(* IEC 61131-3 sources: JingjiangMoonbox/Application/Application/任务列表/TensionTask/张力控制/收放牵/其他, 4 files *)

(* ---- AntiNotch.st ---- *)
(*@CES
Name=AntiNotch
Type=FunctionBlock
TypeGuid=6f9dac99-8de1-4efc-8465-68ac443b7d08
Guid=24b15fba-c20e-4805-94ad-f0677bc5936e
HasDeclaration=True
HasImplementation=True
*)
{DECLARATION}
FUNCTION AntiNotch : BOOL
(*功能：反陷波器(s^2+2*d*wn*s+wn^2)/(s^2+2*d*xi*wn*s+wn^2)的差分方程实现*)
(*输入：*)
(*输出：*)
VAR_INPUT
	i_rU:REAL;(*信号输入*)
	i_prYout: POINTER TO REAL;(*信号输出*)

(*(s^2+2*d*wn*s+wn^2)/(s^2+2*d*xi*wn*s+wn^2)*)
	i_rWn:REAL;(*陷波中心频率 rad/s*)
	i_rBw:REAL;(*陷波宽度 rad/s*)
	i_rDp:REAL;(*陷波深度 dB*)

	i_rTs:REAL;(*采样时间*)

	i_prUk:POINTER TO ARRAY [1..3] OF REAL;(*输入寄存器*)
	i_prYk:POINTER TO ARRAY [1..3] OF REAL;(*输出寄存器*)
END_VAR
VAR
	rFn:REAL:=0;
	rFBw:REAL:=0;
	rWn:REAL:=0;
	rDp:REAL:=0;

	rD:REAL:=0;
	rXi:REAL:=0;

	rK:REAL:=0;
	ra2:REAL:=0;
	ra1:REAL:=0;
	ra0:REAL:=0;

	rb2:REAL:=0;
	rb1:REAL:=0;
	rb0:REAL:=0;

	rTs:REAL:=0;(*采样时间*)
	rTemp:REAL:=0;

END_VAR
{IMPLEMENTATION}
(*参数初始化*)
rFn := LREAL_TO_REAL(i_rWn/2.0*gc_lrPi);
rWn := i_rWn;
rFBw := LREAL_TO_REAL(i_rBw/2.0*gc_lrPi);
rDp := i_rDp;

rTemp := -rDp/20.0;
rD := LREAL_TO_REAL(EXPT(10,rTemp));

rTemp := LREAL_TO_REAL(1.0/(1.0 - 2.0*EXPT(rD,2)));
rXi := rFBw/(2.0*rFn)*SQRT(rTemp);

rK := 1.0;

ra2:=1.0;
ra1:=2*rXi*rWn;
ra0:=rWn*rWn;

rb2:=1;
rb1:=2*rD*rXi*rWn;
rb0:=rWn*rWn;

rTs:=i_rTs;

(*更新寄存器注意顺序*)
i_prYk^[3]:=i_prYk^[2];
i_prYk^[2]:=i_prYk^[1];

i_prUk^[3]:=i_prUk^[2];
i_prUk^[2]:=i_prUk^[1];

(*差分计算*)
i_prUk^[1]:=rK*i_rU;
rTemp:=1/(rb0*rTs*rTs+2*rb1*rTs+4*rb2)*(-(2*rb0*rTs*rTs-8*rb2)*i_prYk^[2]-(rb0*rTs*rTs-2*rb1*rTs+4*rb2)*i_prYk^[3]
            +(ra0*rTs*rTs+2*ra1*rTs+4*ra2)*i_prUk^[1]+(2*ra0*rTs*rTs-8*ra2)*i_prUk^[2]+(ra0*rTs*rTs-2*ra1*rTs+4*ra2)*i_prUk^[3]);
i_prYk^[1]:=rTemp;
i_prYout^:=rTemp;

(* ---- KS_A2B_SmoothDeal.st ---- *)
(*@CES
Name=KS_A2B_SmoothDeal
Type=FunctionBlock
TypeGuid=6f9dac99-8de1-4efc-8465-68ac443b7d08
Guid=9cfb7a1c-ce6a-4c3a-85a6-d0a941a33b90
HasDeclaration=True
HasImplementation=True
*)
{DECLARATION}
FUNCTION KS_A2B_SmoothDeal : REAL
(*从A变化到B平滑处理,返回当前值*)
VAR_INPUT
	i_rA:REAL;
	i_rB:REAL;
	i_rDelta:REAL;(*变化值*)
END_VAR
VAR
	rC:REAL;
END_VAR
{IMPLEMENTATION}
IF i_rDelta<>0 THEN
	IF i_rA > i_rB THEN
		rC:= i_rA - i_rDelta;
		IF rC < i_rB THEN(*限值处理*)
			rC:=i_rB;
		END_IF
	ELSIF i_rA < i_rB THEN
		rC:= i_rA + i_rDelta;
		IF rC > i_rB THEN(*限值处理*)
			rC:=i_rB;
		END_IF
	ELSE
		rC:= i_rB;
	END_IF
ELSE
	rC:=i_rB;
END_IF

KS_A2B_SmoothDeal:=rC;

(* ---- KS_SIG_SIN.st ---- *)
(*@CES
Name=KS_SIG_SIN
Type=FunctionBlock
TypeGuid=6f9dac99-8de1-4efc-8465-68ac443b7d08
Guid=c56967f0-af3c-4951-929b-0432ccffd3b8
HasDeclaration=True
HasImplementation=True
*)
{DECLARATION}
FUNCTION KS_SIG_SIN : BOOL
(*正弦信号*)
VAR_INPUT
	i_xEn:BOOL;(*使能*)
	i_rFreq:REAL;(*频率@hz*)
	i_rAmplitude:REAL;(*幅值*)
	i_uiTotalTime:UINT;(*输出的总时间|=0 代表一直输出@s*)
	i_iCycleTime_Plc:INT;(*程序时间@ms*)
	i_pxOuting:POINTER TO BOOL;(*输出中@如果取消使能,停止到0时结束*)
	i_plrX:POINTER TO LREAL;(*X轴的值*)
	i_prResult:POINTER TO REAL;(*结果值*)
END_VAR
VAR
	xOuting:BOOL;
	lrX:LREAL;(*x值*)
	rResult: REAL;
	lrW:LREAL;(*角速度@rad/s*)
	lrpi: LREAL := 3.1415926;(*圆周率*)
	lrTs: LREAL;(*周期@s*)
	lrTmp: LREAL;
	lrTotalTime:LREAL;(*输出的总时间@ms*)
	xStopOuting: BOOL;
END_VAR
{IMPLEMENTATION}
IF i_rFreq<>0 AND i_rAmplitude<>0 AND i_iCycleTime_Plc<>0 THEN;
ELSE
	RETURN;
END_IF

IF i_pxOuting<>0 THEN
	xOuting:=i_pxOuting^;
END_IF
IF i_plrX<>0 THEN
	lrX:=i_plrX^;
END_IF
IF i_prResult<>0 THEN
	rResult:=i_prResult^;
END_IF

(*使能*)
IF i_xEn THEN
	IF NOT xOuting AND
		lrX = 0 THEN(*lrx用来控制区分是使能取消还是输出完成使用@取消使能才清零*)
		xOuting:=TRUE;
		lrX:=0;(*从0开始*)
	END_IF
END_IF

lrW:=2*lrpi*i_rFreq;(*rad/s*)
lrTs:=1/i_rFreq;(*周期@s*)
lrTotalTime:=UINT_TO_LREAL(i_uiTotalTime)*1000;
IF xOuting THEN
	lrTmp:=lrX / 1000.0;(*s*)
(*
	IF lrTmp>lrTs THEN(*过周期@拉回到一个周期内防止溢出*)
		lrTmp:=lrTmp-lrTs;
	END_IF
*)
	rResult:=LREAL_TO_REAL(i_rAmplitude*SIN(lrW*lrTmp));

	(*更新*)
	xStopOuting:=FALSE;
	IF lrTotalTime<>0 THEN
		IF lrX>=lrTotalTime THEN(*超过了输出的时间*)
			xStopOuting:=TRUE;(*停止输出了*)
		END_IF
	ELSE(*一直输出*);
	END_IF

	lrX:=lrX + i_iCycleTime_Plc;(*ms@也是有可能溢出的|按照pt的经验 先不考虑*)

	IF NOT i_xEn OR xStopOuting THEN(*停止使能\或者停止输出*)
		IF rResult*i_prResult^<=0 THEN(*过零*)
			xOuting:=FALSE;
			rResult:=0;
		END_IF
	END_IF
ELSE
	(*lrx用来控制区分是使能取消还是输出完成使用@取消使能才清零*)
	IF NOT i_xEn THEN
		lrX:=0;
	END_IF
	rResult:=0;
END_IF

IF i_pxOuting<>0 THEN
	i_pxOuting^:=xOuting;
END_IF
IF i_plrX<>0 THEN
	i_plrX^:=lrX;
END_IF
IF i_prResult<>0 THEN
	i_prResult^:=rResult;
END_IF

(* ---- PID_ANTI.st ---- *)
(*@CES
Name=PID_ANTI
Type=FunctionBlock
TypeGuid=6f9dac99-8de1-4efc-8465-68ac443b7d08
Guid=ddf7a214-0c45-4257-a0f0-8ae2d0e2601d
HasDeclaration=True
HasImplementation=True
*)
{DECLARATION}
FUNCTION PID_ANTI : BOOL
VAR_INPUT
(*输入输出*)
	i_rU:REAL;(*控制器输入*)
	i_prYout: POINTER TO REAL;(*控制器输出@绝对值输出*)
(*PID参数*)
	i_rP:REAL;
	i_rI:REAL;
	i_rD:REAL;
	i_rN:REAL;
	i_rTs:REAL;(*s*)
(*积分抗饱和*)
	i_rLim:REAL;(*控制器输出限幅*)
	i_rAntiWindup:REAL;(*抗积分饱和系数@0-->1*)
(*寄存器*)
	i_prYI: POINTER TO REAL;(*积分控制输出寄存器*)
	i_prYD: POINTER TO REAL;(*微分控制输出寄存器*)
	i_parEk:POINTER TO ARRAY [1..2] OF REAL;(*误差寄存器 [e(k);e(k-1)]*)
END_VAR
VAR
	rP:REAL;(*比例部分*)
	rI:REAL;(*积分部分*)
	rD:REAL:=0;(*微分部分*)

	rUnsat:REAL;(*未限幅输出*)
	rTs:REAL:=0;

END_VAR
{IMPLEMENTATION}
(*计算采样时间*)
rTs := i_rTs;

(*误差寄存器更新*)
i_parEk^[2] := i_parEk^[1];
i_parEk^[1] := i_rU;

(*计算比例部分*)
rP := i_rP*i_rU;

(*计算积分部分*)
rI := i_prYI^ + i_rI*i_rU*rTs;
(*计算微分*)
rD := i_prYD^ * (1.0 - i_rN * rTs) + i_rD * i_rN * (i_parEk^[1] - i_parEk^[2]);

(*计算未限幅输出*)
rUnsat := rP + rI + rD;

(*抗积分饱和*)
IF rUnsat>i_rLim THEN
	i_prYout^ := i_rLim;
	rI:=rI - i_rAntiWindup*(rUnsat - i_rLim);
ELSIF rUnsat < -i_rLim THEN
	i_prYout^ := -i_rLim;
	rI:=rI - i_rAntiWindup*(rUnsat + i_rLim);
ELSE
	i_prYout^ := rUnsat;
END_IF

(*寄存器更新*)
i_prYI^ := rI;
i_prYD^ := rD;
